	                //CNV 2
	                IF ("Control_DB".ECnv_Sys[#i_Sys].Instruction.Inbound_Ready OR "Settings_DB".LCnv_Sys[#i_Sys].Cnv_Level[#i_Lev].Cnv2.Cnv_Level = 1) AND
	                    ("Control_DB".VTD_Sys[#i_Sys].Current_Level = #i_Lev OR "Settings_DB".LCnv_Sys[#i_Sys].Cnv_Level[#i_Lev].Cnv2.Cnv_Level = 1) AND
	                    (NOT "Control_DB".LCnv_Sys[#i_Sys].Cnv_Level[#i_Lev].Cnv1.Instruction.Transfer_in_Progress OR "Settings_DB".LCnv_Sys[#i_Sys].Cnv_Level[#i_Lev].Cnv2.Cnv_Level = 1) AND
	                    "Control_DB".LCnv_Sys[#i_Sys].Cnv_Level[#i_Lev].Cnv2.Cnv_Occupied AND
	                    NOT "Control_DB".LCnv_Sys[#i_Sys].Cnv_Level[#i_Lev].Cnv2.Error AND NOT "Control_DB".LCnv_Sys[#i_Sys].Cnv_Level[#i_Lev].Cnv2.Running AND
	                    ("Control_DB".LCnv_Sys[#i_Sys].Cnv_Level[#i_Lev].Cnv2.Mode = 2 OR "Control_DB".LCnv_Sys[#i_Sys].Cnv_Level[#i_Lev].Cnv2.Mode = 3) THEN
	                    "Control_DB".LCnv_Sys[#i_Sys].Cnv_Level[#i_Lev].Cnv2.Instruction.Outbound_Ready := TRUE;
	                ELSIF  NOT "Control_DB".LCnv_Sys[#i_Sys].Cnv_Level[#i_Lev].Cnv2.Cnv_Occupied THEN  // // // // // // // // // // // // //last change
	                    "Control_DB".LCnv_Sys[#i_Sys].Cnv_Level[#i_Lev].Cnv2.Instruction.Outbound_Ready := FALSE;  // // // // // // // // // // // // //last change
	                END_IF;
	            END_FOR;
	        END_REGION

	        REGION TRANSFER IN PROGRESS FOR EXTRACTOR CONVEYOR
	            FOR #i_Lev := "Settings_DB".VTD_Sys[#i_Sys].Lowest_Level TO "Settings_DB".VTD_Sys[#i_Sys].Highest_Level DO
	                "Control_DB".ECnv_Sys[#i_Sys].Instruction.Transfer_in_Progress :=
	                ("Settings_DB".ECnv_Sys[#i_Sys].Cnv_Level = #i_Lev AND
	                "Control_DB".LCnv_Sys[#i_Sys].Cnv_Level[#i_Lev].Cnv1.Instruction.Transfer_in_Progress OR "Control_DB".LCnv_Sys[#i_Sys].Cnv_Level[#i_Lev].Cnv2.Instruction.Transfer_in_Progress);
	            END_FOR;
	        END_REGION
	    END_FOR;

	    IF "FirstScan" THEN
	        "Time_1_Start_Buffers" := T#500MS;
	        "Time_1_end_Buffers" := T#1S;
	        "Time_2_Start_Buffers" := T#1S;
	        "Time_2_End_Buffers" := T#1S_500MS;
	        "Time_3_Buffers" := T#1S_500MS;

	        "Time_1_Start_Ecnv" := T#1S_700MS;
	        "Time_1_end_Ecnv" := T#2S_100MS;
	        "Time_2_Start_Ecnv" := T#2S_100MS;
	        "Time_2_End_Ecnv" := T#2S_600MS;
	        "Time_3_Ecnv" := T#2S_600MS;
	    END_IF;


END_FUNCTION

